(* IEC 61131-3 sources: MHFW-01/plc/function_blocks, 11 files *)

(* ---- FB_AlarmManager.st ---- *)
FUNCTION_BLOCK FB_AlarmManager
VAR_INPUT
  Cause : INT;
  ResetPB : BOOL;
  RecoveryOK : BOOL;
  Cold : BOOL;
END_VAR
VAR_OUTPUT
  Alarm : INT;
END_VAR
VAR
  PrevReset : BOOL;
END_VAR
IF Cold THEN Alarm := 0; END_IF;
IF ResetPB AND NOT PrevReset AND RecoveryOK THEN Alarm := 0; END_IF;
IF Cause <> 0 THEN Alarm := Cause; END_IF;
PrevReset := ResetPB;
END_FUNCTION_BLOCK

(* ---- FB_AxisSynchronization.st ---- *)
FUNCTION_BLOCK FB_AxisSynchronization
VAR_INPUT
  Phase : REAL;
  Offset : REAL;
END_VAR
VAR_OUTPUT
  SealPhase : REAL;
  JawTarget : REAL;
  Close : BOOL;
END_VAR
VAR
  Distance : REAL;
END_VAR
SealPhase := Phase + Offset;
SealPhase := SealPhase - DINT_TO_REAL(TRUNC(SealPhase));
IF SealPhase < 0.0 THEN SealPhase := SealPhase + 1.0; END_IF;
Distance := MIN(SealPhase, 1.0 - SealPhase);
(* Electronic cam: closed dwell +/-0.04, ramp to fully open at 0.20. *)
JawTarget := LIMIT(0.0, (Distance - 0.04) * 250.0, 40.0);
Close := Distance < 0.04;
END_FUNCTION_BLOCK

(* ---- FB_BagLengthControl.st ---- *)
FUNCTION_BLOCK FB_BagLengthControl
VAR_INPUT
  Position : REAL;
  Pitch : REAL;
  Offset : REAL;
  Reset : BOOL;
END_VAR
VAR_OUTPUT
  Phase : REAL;
  Boundary : BOOL;
END_VAR
VAR
  Previous : REAL;
  Turns : REAL;
END_VAR
Turns := (Position + Offset) / Pitch;
Phase := Turns - DINT_TO_REAL(TRUNC(Turns));
IF Phase < 0.0 THEN Phase := Phase + 1.0; END_IF;
Boundary := (Phase < Previous) AND NOT Reset;
Previous := Phase;
END_FUNCTION_BLOCK

(* ---- FB_CenterSeal.st ---- *)
FUNCTION_BLOCK FB_CenterSeal
VAR_INPUT
  Enable : BOOL;
  Fresh : BOOL;
  Reset : BOOL;
  Speed : REAL;
  StepSeconds : REAL;
END_VAR
VAR_OUTPUT
  Run : BOOL;
  Target : REAL;
END_VAR
VAR
END_VAR
IF Reset THEN Target := 0.0; END_IF;
Run := Enable;
IF Enable AND Fresh THEN Target := Target + Speed * StepSeconds; END_IF;
END_FUNCTION_BLOCK

(* ---- FB_Cutter.st ---- *)
FUNCTION_BLOCK FB_Cutter
VAR_INPUT
  Enable : BOOL;
  Boundary : BOOL;
  SealClose : BOOL;
END_VAR
VAR_OUTPUT
  Pulse : BOOL;
END_VAR
VAR
END_VAR
Pulse := Enable AND Boundary AND SealClose;
END_FUNCTION_BLOCK

(* ---- FB_Discharge.st ---- *)
FUNCTION_BLOCK FB_Discharge
VAR_INPUT
  Enable : BOOL;
  Fresh : BOOL;
  Reset : BOOL;
  Speed : REAL;
  StepSeconds : REAL;
END_VAR
VAR_OUTPUT
  Run : BOOL;
  Target : REAL;
END_VAR
VAR
END_VAR
IF Reset THEN Target := 0.0; END_IF;
Run := Enable;
IF Enable AND Fresh THEN Target := Target + Speed * StepSeconds; END_IF;
END_FUNCTION_BLOCK

(* ---- FB_EndSeal.st ---- *)
FUNCTION_BLOCK FB_EndSeal
VAR_INPUT
  Enable : BOOL;
  CamClose : BOOL;
  CamTarget : REAL;
END_VAR
VAR_OUTPUT
  Close : BOOL;
  Target : REAL;
END_VAR
VAR
END_VAR
Close := Enable AND CamClose;
IF Enable THEN Target := CamTarget; ELSE Target := 40.0; END_IF;
END_FUNCTION_BLOCK

(* ---- FB_FilmFeed.st ---- *)
FUNCTION_BLOCK FB_FilmFeed
VAR_INPUT
  Enable : BOOL;
  Fresh : BOOL;
  Reset : BOOL;
  Speed : REAL;
  StepSeconds : REAL;
END_VAR
VAR_OUTPUT
  Run : BOOL;
  Target : REAL;
END_VAR
VAR
END_VAR
IF Reset THEN Target := 0.0; END_IF;
Run := Enable;
IF Enable AND Fresh THEN Target := Target + Speed * StepSeconds; END_IF;
END_FUNCTION_BLOCK

(* ---- FB_InfeedConveyor.st ---- *)
FUNCTION_BLOCK FB_InfeedConveyor
VAR_INPUT
  Enable : BOOL;
  Fresh : BOOL;
  Reset : BOOL;
  Speed : REAL;
  StepSeconds : REAL;
END_VAR
VAR_OUTPUT
  Run : BOOL;
  Target : REAL;
END_VAR
VAR
END_VAR
IF Reset THEN Target := 0.0; END_IF;
Run := Enable;
IF Enable AND Fresh THEN Target := Target + Speed * StepSeconds; END_IF;
END_FUNCTION_BLOCK

(* ---- FB_ModeManager.st ---- *)
FUNCTION_BLOCK FB_ModeManager
VAR_INPUT
  StartPB : BOOL;
  StopPB : BOOL;
  Requested : INT;
  Alarm : INT;
  SingleDone : BOOL;
  Cold : BOOL;
END_VAR
VAR_OUTPUT
  Running : BOOL;
  Mode : INT;
END_VAR
VAR
  PrevStart : BOOL;
END_VAR
IF Cold THEN Running := FALSE; Mode := 4; END_IF;
IF Alarm = 0 AND Mode = 5 THEN Mode := 4; END_IF;
IF StartPB AND NOT PrevStart AND Alarm = 0 AND Requested >= 1 AND Requested <= 3 THEN Running := TRUE; Mode := Requested; END_IF;
IF StopPB OR SingleDone THEN Running := FALSE; Mode := 4; END_IF;
IF Alarm <> 0 THEN Running := FALSE; Mode := 5; END_IF;
PrevStart := StartPB;
END_FUNCTION_BLOCK

(* ---- FB_ProductDetection.st ---- *)
FUNCTION_BLOCK FB_ProductDetection
VAR_INPUT
  Present : BOOL;
  Run : BOOL;
  Fresh : BOOL;
  StepSeconds : REAL;
  Period : REAL;
  Reset : BOOL;
END_VAR
VAR_OUTPUT
  Missing : BOOL;
  StuckOn : BOOL;
END_VAR
VAR
  AbsentTime : REAL;
  PresentTime : REAL;
END_VAR
IF Reset OR NOT Run THEN AbsentTime := 0.0; PresentTime := 0.0; END_IF;
IF Run AND Fresh THEN
 IF Present THEN AbsentTime := 0.0; PresentTime := PresentTime + StepSeconds;
 ELSE PresentTime := 0.0; AbsentTime := AbsentTime + StepSeconds; END_IF;
END_IF;
Missing := AbsentTime > 2.2 * Period;
StuckOn := PresentTime > 1.2 * Period;
END_FUNCTION_BLOCK
